Fanuc KAREL source: kx00015.KL

-- PROVISIONAL review KL for V940-1; original PC SHA256 8b5443bdf8feaa8ac2cf91ca3a1ea57cfbb772087b631a6612e83d93be49bbcd
-- Incomplete behavior may be omitted. Consult companion uncertainty JSON. Do not deploy.
PROGRAM KX00015
%NOLOCKGROUP
VAR
  I : INTEGER
  J : INTEGER
  B : BOOLEAN
  F : FILE
  S : STRING[80]
-- UNRESOLVED_DECL P type=000102
BEGIN
  -- V9_ZERO_TABLE_METADATA_HINT layout=0001; no indexed target words; source/name/runtime held
  -- UNRESOLVED_PC offsets 5-7; opcodes 9D,0E
  -- UNRESOLVED_PC offsets 12-16; opcodes 7F
END KX00015
